Fanuc KAREL source: KA00031.KL

PROGRAM KA00031
%NOLOCKGROUP
VAR
  SRC: BOOLEAN
  DST: XYZWPREXT
BEGIN
  SRC = TRUE
  DST = SRC
END KA00031
